(* IEC 61131-3 sources: trust-platform/crates/trust-runtime/tests/fixtures/plcopen_motion/single_axis_core/src (part 2) *)

TEST_PROGRAM plcopen_motion_single_axis_buffer_mode_support_rules_by_fb_family
VAR
    AxisHomeBuffered : AXIS_REF;
    AxisHomeUnsupported : AXIS_REF;
    AxisHaltUnsupported : AXIS_REF;
    AxisAdditiveUnsupported : AXIS_REF;
    AxisVelocityBuffered : AXIS_REF;
    AxisVelocityUnsupported : AXIS_REF;
    AxisContinuousBuffered : AXIS_REF;
    AxisContinuousUnsupported : AXIS_REF;
    SeedHomeBuffered : TRUST_MOTION_TestAxisSeed;
    SeedHomeUnsupported : TRUST_MOTION_TestAxisSeed;
    SeedHaltUnsupported : TRUST_MOTION_TestAxisSeed;
    SeedAdditiveUnsupported : TRUST_MOTION_TestAxisSeed;
    SeedVelocityBuffered : TRUST_MOTION_TestAxisSeed;
    SeedVelocityUnsupported : TRUST_MOTION_TestAxisSeed;
    SeedContinuousBuffered : TRUST_MOTION_TestAxisSeed;
    SeedContinuousUnsupported : TRUST_MOTION_TestAxisSeed;
    HomeBuffered : MC_Home;
    HomeUnsupported : MC_Home;
    HaltUnsupported : MC_Halt;
    MoveAdditiveUnsupported : MC_MoveAdditive;
    MoveVelocityBuffered : MC_MoveVelocity;
    MoveVelocityUnsupported : MC_MoveVelocity;
    MoveContinuousAbsoluteBuffered : MC_MoveContinuousAbsolute;
    MoveContinuousRelativeUnsupported : MC_MoveContinuousRelative;
END_VAR

AxisHomeBuffered.AxisId := UDINT#139;
AxisHomeBuffered.InternalIndex := UINT#18;
SeedHomeBuffered(Axis := AxisHomeBuffered, ResetDefaults := TRUE, ApplyState := TRUE, State := MC_AXIS_STATUS#mcStandstill);
HomeBuffered(Axis := AxisHomeBuffered, Execute := TRUE, Position := REAL#5.0, BufferMode := MC_BUFFER_MODE#mcBuffered);
ASSERT_TRUE(HomeBuffered.Busy);
ASSERT_TRUE(HomeBuffered.Active);
ASSERT_FALSE(HomeBuffered.Error);

AxisHomeUnsupported.AxisId := UDINT#140;
AxisHomeUnsupported.InternalIndex := UINT#19;
SeedHomeUnsupported(Axis := AxisHomeUnsupported, ResetDefaults := TRUE, ApplyState := TRUE, State := MC_AXIS_STATUS#mcStandstill);
HomeUnsupported(Axis := AxisHomeUnsupported, Execute := TRUE, Position := REAL#5.0, BufferMode := MC_BUFFER_MODE#mcBlendingLow);
ASSERT_TRUE(HomeUnsupported.Error);
ASSERT_TRUE(HomeUnsupported.ErrorID = WORD#16#0500);

AxisHaltUnsupported.AxisId := UDINT#141;
AxisHaltUnsupported.InternalIndex := UINT#20;
SeedHaltUnsupported(Axis := AxisHaltUnsupported, ResetDefaults := TRUE, ApplyState := TRUE, State := MC_AXIS_STATUS#mcContinuousMotion);
HaltUnsupported(Axis := AxisHaltUnsupported, Execute := TRUE, Deceleration := REAL#2.0, Jerk := REAL#1.0, BufferMode := MC_BUFFER_MODE#mcBlendingLow);
ASSERT_TRUE(HaltUnsupported.Error);
ASSERT_TRUE(HaltUnsupported.ErrorID = WORD#16#0500);

AxisAdditiveUnsupported.AxisId := UDINT#142;
AxisAdditiveUnsupported.InternalIndex := UINT#21;
SeedAdditiveUnsupported(
    Axis := AxisAdditiveUnsupported,
    ResetDefaults := TRUE,
    ApplyState := TRUE,
    State := MC_AXIS_STATUS#mcStandstill,
    ApplyActuals := TRUE,
    ActualPosition := REAL#10.0,
    SetPosition := REAL#10.0,
    CommandedPosition := REAL#10.0,
    ActualVelocity := REAL#0.0,
    SetVelocity := REAL#0.0,
    CommandedVelocity := REAL#0.0,
    ActualTorque := REAL#0.0
);
MoveAdditiveUnsupported(Axis := AxisAdditiveUnsupported, Execute := TRUE, ContinuousUpdate := FALSE, Distance := REAL#5.0, Velocity := REAL#4.0, Acceleration := REAL#2.0, Deceleration := REAL#2.0, Jerk := REAL#1.0, BufferMode := MC_BUFFER_MODE#mcBlendingLow);
ASSERT_TRUE(MoveAdditiveUnsupported.Error);
ASSERT_TRUE(MoveAdditiveUnsupported.ErrorID = WORD#16#0500);

AxisVelocityBuffered.AxisId := UDINT#143;
AxisVelocityBuffered.InternalIndex := UINT#22;
SeedVelocityBuffered(Axis := AxisVelocityBuffered, ResetDefaults := TRUE, ApplyState := TRUE, State := MC_AXIS_STATUS#mcStandstill);
MoveVelocityBuffered(Axis := AxisVelocityBuffered, Execute := TRUE, ContinuousUpdate := FALSE, Velocity := REAL#4.0, Acceleration := REAL#2.0, Deceleration := REAL#2.0, Jerk := REAL#1.0, Direction := MC_DIRECTION#mcCurrentDirection, BufferMode := MC_BUFFER_MODE#mcBuffered);
ASSERT_TRUE(MoveVelocityBuffered.Busy);
ASSERT_TRUE(MoveVelocityBuffered.Active);
ASSERT_TRUE(MoveVelocityBuffered.InVelocity);
ASSERT_FALSE(MoveVelocityBuffered.Error);

AxisVelocityUnsupported.AxisId := UDINT#144;
AxisVelocityUnsupported.InternalIndex := UINT#23;
SeedVelocityUnsupported(Axis := AxisVelocityUnsupported, ResetDefaults := TRUE, ApplyState := TRUE, State := MC_AXIS_STATUS#mcStandstill);
MoveVelocityUnsupported(Axis := AxisVelocityUnsupported, Execute := TRUE, ContinuousUpdate := FALSE, Velocity := REAL#4.0, Acceleration := REAL#2.0, Deceleration := REAL#2.0, Jerk := REAL#1.0, Direction := MC_DIRECTION#mcCurrentDirection, BufferMode := MC_BUFFER_MODE#mcBlendingLow);
ASSERT_TRUE(MoveVelocityUnsupported.Error);
ASSERT_TRUE(MoveVelocityUnsupported.ErrorID = WORD#16#0500);

AxisContinuousBuffered.AxisId := UDINT#145;
AxisContinuousBuffered.InternalIndex := UINT#24;
SeedContinuousBuffered(Axis := AxisContinuousBuffered, ResetDefaults := TRUE, ApplyState := TRUE, State := MC_AXIS_STATUS#mcStandstill);
MoveContinuousAbsoluteBuffered(Axis := AxisContinuousBuffered, Execute := TRUE, ContinuousUpdate := FALSE, Position := REAL#30.0, EndVelocity := REAL#3.0, Velocity := REAL#8.0, Acceleration := REAL#4.0, Deceleration := REAL#4.0, Jerk := REAL#1.0, Direction := MC_DIRECTION#mcCurrentDirection, BufferMode := MC_BUFFER_MODE#mcBuffered);
ASSERT_TRUE(MoveContinuousAbsoluteBuffered.Busy);
ASSERT_TRUE(MoveContinuousAbsoluteBuffered.Active);
ASSERT_TRUE(MoveContinuousAbsoluteBuffered.InEndVelocity);
ASSERT_FALSE(MoveContinuousAbsoluteBuffered.Error);

AxisContinuousUnsupported.AxisId := UDINT#146;
AxisContinuousUnsupported.InternalIndex := UINT#25;
SeedContinuousUnsupported(Axis := AxisContinuousUnsupported, ResetDefaults := TRUE, ApplyState := TRUE, State := MC_AXIS_STATUS#mcStandstill);
MoveContinuousRelativeUnsupported(Axis := AxisContinuousUnsupported, Execute := TRUE, ContinuousUpdate := FALSE, Distance := REAL#5.0, EndVelocity := REAL#3.0, Velocity := REAL#8.0, Acceleration := REAL#4.0, Deceleration := REAL#4.0, Jerk := REAL#1.0, BufferMode := MC_BUFFER_MODE#mcBlendingLow);
ASSERT_TRUE(MoveContinuousRelativeUnsupported.Error);
ASSERT_TRUE(MoveContinuousRelativeUnsupported.ErrorID = WORD#16#0500);
END_TEST_PROGRAM

TEST_PROGRAM plcopen_motion_single_axis_home_halt_stop_and_continuous_end_velocity_behaviors
VAR
    AxisHome : AXIS_REF;
    AxisHalt : AXIS_REF;
    AxisStop : AXIS_REF;
    AxisContinuous : AXIS_REF;
    SeedHome : TRUST_MOTION_TestAxisSeed;
    SeedHalt : TRUST_MOTION_TestAxisSeed;
    SeedStop : TRUST_MOTION_TestAxisSeed;
    SeedContinuous : TRUST_MOTION_TestAxisSeed;
    Home : MC_Home;
    Halt : MC_Halt;
    Stop : MC_Stop;
    MoveContinuousAbsolute : MC_MoveContinuousAbsolute;
    ReadStatusHome : MC_ReadStatus;
    ReadStatusHalt : MC_ReadStatus;
    ReadStatusStop : MC_ReadStatus;
    ReadStatusContinuous : MC_ReadStatus;
    ReadAxisInfo : MC_ReadAxisInfo;
    ReadActualVelocity : MC_ReadActualVelocity;
END_VAR

AxisHome.AxisId := UDINT#121;
AxisHome.InternalIndex := UINT#25;
SeedHome(Axis := AxisHome, ResetDefaults := TRUE, ApplyState := TRUE, State := MC_AXIS_STATUS#mcStandstill, ApplyPowerStage := TRUE, PowerStage := TRUE);
Home(Axis := AxisHome, Execute := TRUE, Position := REAL#12.0, BufferMode := MC_BUFFER_MODE#mcAborting);
ASSERT_TRUE(Home.Busy);
ASSERT_TRUE(Home.Active);
ReadStatusHome(Axis := AxisHome, Enable := TRUE);
ASSERT_TRUE(ReadStatusHome.Homing);
Home(Axis := AxisHome, Execute := FALSE, Position := REAL#12.0, BufferMode := MC_BUFFER_MODE#mcAborting);
ASSERT_TRUE(Home.Done);
ReadStatusHome(Axis := AxisHome, Enable := TRUE);
ASSERT_TRUE(ReadStatusHome.Standstill);
ReadAxisInfo(Axis := AxisHome, Enable := TRUE);
ASSERT_TRUE(ReadAxisInfo.IsHomed);

AxisHalt.AxisId := UDINT#122;
AxisHalt.InternalIndex := UINT#26;
SeedHalt(Axis := AxisHalt, ResetDefaults := TRUE, ApplyState := TRUE, State := MC_AXIS_STATUS#mcContinuousMotion, ApplyPowerStage := TRUE, PowerStage := TRUE);
Halt(Axis := AxisHalt, Execute := TRUE, Deceleration := REAL#2.0, Jerk := REAL#1.0, BufferMode := MC_BUFFER_MODE#mcBuffered);
ASSERT_TRUE(Halt.Busy);
ASSERT_TRUE(Halt.Active);
ReadStatusHalt(Axis := AxisHalt, Enable := TRUE);
ASSERT_TRUE(ReadStatusHalt.DiscreteMotion);
ASSERT_FALSE(ReadStatusHalt.Stopping);
Halt(Axis := AxisHalt, Execute := FALSE, Deceleration := REAL#2.0, Jerk := REAL#1.0, BufferMode := MC_BUFFER_MODE#mcBuffered);
ASSERT_TRUE(Halt.Done);
ReadStatusHalt(Axis := AxisHalt, Enable := TRUE);
ASSERT_TRUE(ReadStatusHalt.Standstill);

AxisStop.AxisId := UDINT#123;
AxisStop.InternalIndex := UINT#27;
SeedStop(Axis := AxisStop, ResetDefaults := TRUE, ApplyState := TRUE, State := MC_AXIS_STATUS#mcContinuousMotion, ApplyPowerStage := TRUE, PowerStage := TRUE);
Stop(Axis := AxisStop, Execute := TRUE, Deceleration := REAL#2.0, Jerk := REAL#1.0);
ASSERT_FALSE(Stop.Busy);
ASSERT_TRUE(Stop.Done);
ReadStatusStop(Axis := AxisStop, Enable := TRUE);
ASSERT_TRUE(ReadStatusStop.Stopping);
Stop(Axis := AxisStop, Execute := FALSE, Deceleration := REAL#2.0, Jerk := REAL#1.0);
ASSERT_TRUE(Stop.Done);
ReadStatusStop(Axis := AxisStop, Enable := TRUE);
ASSERT_TRUE(ReadStatusStop.Standstill);

AxisContinuous.AxisId := UDINT#124;
AxisContinuous.InternalIndex := UINT#28;
SeedContinuous(Axis := AxisContinuous, ResetDefaults := TRUE, ApplyState := TRUE, State := MC_AXIS_STATUS#mcStandstill);
MoveContinuousAbsolute(
    Axis := AxisContinuous,
    Execute := TRUE,
    ContinuousUpdate := FALSE,
    Position := REAL#40.0,
    EndVelocity := REAL#3.0,
    Velocity := REAL#8.0,
    Acceleration := REAL#4.0,
    Deceleration := REAL#4.0,
    Jerk := REAL#1.0,
    Direction := MC_DIRECTION#mcCurrentDirection,
    BufferMode := MC_BUFFER_MODE#mcAborting
);
ASSERT_TRUE(MoveContinuousAbsolute.Busy);
ASSERT_TRUE(MoveContinuousAbsolute.Active);
ASSERT_TRUE(MoveContinuousAbsolute.InEndVelocity);
ReadStatusContinuous(Axis := AxisContinuous, Enable := TRUE);
ASSERT_TRUE(ReadStatusContinuous.ContinuousMotion);
ReadActualVelocity(Axis := AxisContinuous, Enable := TRUE);
ASSERT_TRUE(ReadActualVelocity.Velocity = REAL#3.0);
MoveContinuousAbsolute(
    Axis := AxisContinuous,
    Execute := FALSE,
    ContinuousUpdate := FALSE,
    Position := REAL#40.0,
    EndVelocity := REAL#3.0,
    Velocity := REAL#8.0,
    Acceleration := REAL#4.0,
    Deceleration := REAL#4.0,
    Jerk := REAL#1.0,
    Direction := MC_DIRECTION#mcCurrentDirection,
    BufferMode := MC_BUFFER_MODE#mcAborting
);
ASSERT_FALSE(MoveContinuousAbsolute.InEndVelocity);
ReadStatusContinuous(Axis := AxisContinuous, Enable := TRUE);
ASSERT_TRUE(ReadStatusContinuous.Standstill);
END_TEST_PROGRAM

TEST_PROGRAM plcopen_motion_single_axis_continuous_update_changes_target_and_end_velocity
VAR
    AxisAbsolute : AXIS_REF;
    AxisRelative : AXIS_REF;
    SeedAbsolute : TRUST_MOTION_TestAxisSeed;
    SeedRelative : TRUST_MOTION_TestAxisSeed;
    MoveContinuousAbsolute : MC_MoveContinuousAbsolute;
    MoveContinuousRelative : MC_MoveContinuousRelative;
    ReadAbsolute : MC_ReadParameter;
    ReadRelative : MC_ReadParameter;
    ReadVelocityAbsolute : MC_ReadActualVelocity;
    ReadVelocityRelative : MC_ReadActualVelocity;
    Constants : MC_Constants;
END_VAR

Constants();
AxisAbsolute.AxisId := UDINT#147;
AxisAbsolute.InternalIndex := UINT#26;
SeedAbsolute(
    Axis := AxisAbsolute,
    ResetDefaults := TRUE,
    ApplyState := TRUE,
    State := MC_AXIS_STATUS#mcStandstill,
    ApplyActuals := TRUE,
    ActualPosition := REAL#10.0,
    SetPosition := REAL#10.0,
    CommandedPosition := REAL#10.0,
    ActualVelocity := REAL#0.0,
    SetVelocity := REAL#0.0,
    CommandedVelocity := REAL#0.0,
    ActualTorque := REAL#0.0
);
MoveContinuousAbsolute(Axis := AxisAbsolute, Execute := TRUE, ContinuousUpdate := FALSE, Position := REAL#40.0, EndVelocity := REAL#3.0, Velocity := REAL#8.0, Acceleration := REAL#4.0, Deceleration := REAL#4.0, Jerk := REAL#1.0, Direction := MC_DIRECTION#mcCurrentDirection, BufferMode := MC_BUFFER_MODE#mcAborting);
MoveContinuousAbsolute(Axis := AxisAbsolute, Execute := TRUE, ContinuousUpdate := TRUE, Position := REAL#55.0, EndVelocity := REAL#4.0, Velocity := REAL#8.0, Acceleration := REAL#4.0, Deceleration := REAL#4.0, Jerk := REAL#1.0, Direction := MC_DIRECTION#mcCurrentDirection, BufferMode := MC_BUFFER_MODE#mcAborting);
ASSERT_TRUE(MoveContinuousAbsolute.InEndVelocity);
ReadAbsolute(Axis := AxisAbsolute, Enable := TRUE, ParameterNumber := Constants.PN_CommandedPosition);
ASSERT_TRUE(ReadAbsolute.Value = REAL#55.0);
ReadVelocityAbsolute(Axis := AxisAbsolute, Enable := TRUE);
ASSERT_TRUE(ReadVelocityAbsolute.Velocity = REAL#4.0);

AxisRelative.AxisId := UDINT#148;
AxisRelative.InternalIndex := UINT#27;
SeedRelative(
    Axis := AxisRelative,
    ResetDefaults := TRUE,
    ApplyState := TRUE,
    State := MC_AXIS_STATUS#mcStandstill,
    ApplyActuals := TRUE,
    ActualPosition := REAL#10.0,
    SetPosition := REAL#10.0,
    CommandedPosition := REAL#10.0,
    ActualVelocity := REAL#0.0,
    SetVelocity := REAL#0.0,
    CommandedVelocity := REAL#0.0,
    ActualTorque := REAL#0.0
);
MoveContinuousRelative(Axis := AxisRelative, Execute := TRUE, ContinuousUpdate := FALSE, Distance := REAL#5.0, EndVelocity := REAL#2.0, Velocity := REAL#8.0, Acceleration := REAL#4.0, Deceleration := REAL#4.0, Jerk := REAL#1.0, BufferMode := MC_BUFFER_MODE#mcAborting);
MoveContinuousRelative(Axis := AxisRelative, Execute := TRUE, ContinuousUpdate := TRUE, Distance := REAL#8.0, EndVelocity := REAL#4.0, Velocity := REAL#8.0, Acceleration := REAL#4.0, Deceleration := REAL#4.0, Jerk := REAL#1.0, BufferMode := MC_BUFFER_MODE#mcAborting);
ASSERT_TRUE(MoveContinuousRelative.InEndVelocity);
ReadRelative(Axis := AxisRelative, Enable := TRUE, ParameterNumber := Constants.PN_CommandedPosition);
ASSERT_TRUE(ReadRelative.Value = REAL#18.0);
ReadVelocityRelative(Axis := AxisRelative, Enable := TRUE);
ASSERT_TRUE(ReadVelocityRelative.Velocity = REAL#4.0);
END_TEST_PROGRAM

TEST_PROGRAM plcopen_motion_single_axis_continuous_commandaborted_resets_in_end_velocity
VAR
    Axis : AXIS_REF;
    Seed : TRUST_MOTION_TestAxisSeed;
    MoveContinuous : MC_MoveContinuousAbsolute;
    MoveAbort : MC_MoveAbsolute;
    ReadStatus : MC_ReadStatus;
END_VAR

Axis.AxisId := UDINT#149;
Axis.InternalIndex := UINT#28;
Seed(Axis := Axis, ResetDefaults := TRUE, ApplyState := TRUE, State := MC_AXIS_STATUS#mcStandstill);
MoveContinuous(Axis := Axis, Execute := TRUE, ContinuousUpdate := FALSE, Position := REAL#30.0, EndVelocity := REAL#3.0, Velocity := REAL#8.0, Acceleration := REAL#4.0, Deceleration := REAL#4.0, Jerk := REAL#1.0, Direction := MC_DIRECTION#mcCurrentDirection, BufferMode := MC_BUFFER_MODE#mcAborting);
ASSERT_TRUE(MoveContinuous.InEndVelocity);
MoveAbort(Axis := Axis, Execute := TRUE, ContinuousUpdate := FALSE, Position := REAL#12.0, Velocity := REAL#5.0, Acceleration := REAL#2.0, Deceleration := REAL#2.0, Jerk := REAL#1.0, Direction := MC_DIRECTION#mcCurrentDirection, BufferMode := MC_BUFFER_MODE#mcAborting);
ASSERT_TRUE(MoveAbort.Active);
MoveContinuous(Axis := Axis, Execute := TRUE, ContinuousUpdate := FALSE, Position := REAL#30.0, EndVelocity := REAL#3.0, Velocity := REAL#8.0, Acceleration := REAL#4.0, Deceleration := REAL#4.0, Jerk := REAL#1.0, Direction := MC_DIRECTION#mcCurrentDirection, BufferMode := MC_BUFFER_MODE#mcAborting);
ASSERT_TRUE(MoveContinuous.CommandAborted);
ASSERT_FALSE(MoveContinuous.InEndVelocity);
ASSERT_FALSE(MoveContinuous.Busy);
ASSERT_FALSE(MoveContinuous.Active);
ReadStatus(Axis := Axis, Enable := TRUE);
ASSERT_TRUE(ReadStatus.DiscreteMotion);
END_TEST_PROGRAM

TEST_PROGRAM plcopen_motion_single_axis_buffered_home_halt_and_additive_take_ownership_after_active_motion
VAR
    AxisHome : AXIS_REF;
    AxisHalt : AXIS_REF;
    AxisAdditive : AXIS_REF;
    SeedHome : TRUST_MOTION_TestAxisSeed;
    SeedHalt : TRUST_MOTION_TestAxisSeed;
    SeedAdditive : TRUST_MOTION_TestAxisSeed;
    MoveActiveHome : MC_MoveAbsolute;
    MoveActiveHalt : MC_MoveAbsolute;
    MoveActiveAdditive : MC_MoveAbsolute;
    Home : MC_Home;
    Halt : MC_Halt;
    MoveAdditive : MC_MoveAdditive;
    ReadStatusHome : MC_ReadStatus;
    ReadStatusHalt : MC_ReadStatus;
    ReadAxisInfoHome : MC_ReadAxisInfo;
    ReadActualAdditive : MC_ReadActualPosition;
END_VAR

AxisHome.AxisId := UDINT#150;
AxisHome.InternalIndex := UINT#29;
SeedHome(Axis := AxisHome, ResetDefaults := TRUE, ApplyState := TRUE, State := MC_AXIS_STATUS#mcStandstill);
MoveActiveHome(Axis := AxisHome, Execute := TRUE, ContinuousUpdate := FALSE, Position := REAL#15.0, Velocity := REAL#5.0, Acceleration := REAL#2.0, Deceleration := REAL#2.0, Jerk := REAL#1.0, Direction := MC_DIRECTION#mcCurrentDirection, BufferMode := MC_BUFFER_MODE#mcAborting);
Home(Axis := AxisHome, Execute := TRUE, Position := REAL#7.0, BufferMode := MC_BUFFER_MODE#mcBuffered);
ASSERT_TRUE(Home.Busy);
ASSERT_FALSE(Home.Active);
MoveActiveHome(Axis := AxisHome, Execute := FALSE, ContinuousUpdate := FALSE, Position := REAL#15.0, Velocity := REAL#5.0, Acceleration := REAL#2.0, Deceleration := REAL#2.0, Jerk := REAL#1.0, Direction := MC_DIRECTION#mcCurrentDirection, BufferMode := MC_BUFFER_MODE#mcAborting);
Home(Axis := AxisHome, Execute := TRUE, Position := REAL#7.0, BufferMode := MC_BUFFER_MODE#mcBuffered);
ASSERT_TRUE(Home.Active);
ReadStatusHome(Axis := AxisHome, Enable := TRUE);
ASSERT_TRUE(ReadStatusHome.Homing);
Home(Axis := AxisHome, Execute := FALSE, Position := REAL#7.0, BufferMode := MC_BUFFER_MODE#mcBuffered);
ASSERT_TRUE(Home.Done);
ReadAxisInfoHome(Axis := AxisHome, Enable := TRUE);
ASSERT_TRUE(ReadAxisInfoHome.IsHomed);

AxisHalt.AxisId := UDINT#151;
AxisHalt.InternalIndex := UINT#30;
SeedHalt(Axis := AxisHalt, ResetDefaults := TRUE, ApplyState := TRUE, State := MC_AXIS_STATUS#mcStandstill);
MoveActiveHalt(Axis := AxisHalt, Execute := TRUE, ContinuousUpdate := FALSE, Position := REAL#20.0, Velocity := REAL#5.0, Acceleration := REAL#2.0, Deceleration := REAL#2.0, Jerk := REAL#1.0, Direction := MC_DIRECTION#mcCurrentDirection, BufferMode := MC_BUFFER_MODE#mcAborting);
Halt(Axis := AxisHalt, Execute := TRUE, Deceleration := REAL#2.0, Jerk := REAL#1.0, BufferMode := MC_BUFFER_MODE#mcBuffered);
ASSERT_TRUE(Halt.Busy);
ASSERT_FALSE(Halt.Active);
MoveActiveHalt(Axis := AxisHalt, Execute := FALSE, ContinuousUpdate := FALSE, Position := REAL#20.0, Velocity := REAL#5.0, Acceleration := REAL#2.0, Deceleration := REAL#2.0, Jerk := REAL#1.0, Direction := MC_DIRECTION#mcCurrentDirection, BufferMode := MC_BUFFER_MODE#mcAborting);
Halt(Axis := AxisHalt, Execute := TRUE, Deceleration := REAL#2.0, Jerk := REAL#1.0, BufferMode := MC_BUFFER_MODE#mcBuffered);
ASSERT_TRUE(Halt.Active);
ReadStatusHalt(Axis := AxisHalt, Enable := TRUE);
ASSERT_TRUE(ReadStatusHalt.DiscreteMotion);
Halt(Axis := AxisHalt, Execute := FALSE, Deceleration := REAL#2.0, Jerk := REAL#1.0, BufferMode := MC_BUFFER_MODE#mcBuffered);
ASSERT_TRUE(Halt.Done);
ReadStatusHalt(Axis := AxisHalt, Enable := TRUE);
ASSERT_TRUE(ReadStatusHalt.Standstill);

AxisAdditive.AxisId := UDINT#152;
AxisAdditive.InternalIndex := UINT#31;
SeedAdditive(
    Axis := AxisAdditive,
    ResetDefaults := TRUE,
    ApplyState := TRUE,
    State := MC_AXIS_STATUS#mcStandstill,
    ApplyActuals := TRUE,
    ActualPosition := REAL#10.0,
    SetPosition := REAL#10.0,
    CommandedPosition := REAL#10.0,
    ActualVelocity := REAL#0.0,
    SetVelocity := REAL#0.0,
    CommandedVelocity := REAL#0.0,
    ActualTorque := REAL#0.0
);
MoveActiveAdditive(Axis := AxisAdditive, Execute := TRUE, ContinuousUpdate := FALSE, Position := REAL#15.0, Velocity := REAL#5.0, Acceleration := REAL#2.0, Deceleration := REAL#2.0, Jerk := REAL#1.0, Direction := MC_DIRECTION#mcCurrentDirection, BufferMode := MC_BUFFER_MODE#mcAborting);
MoveAdditive(Axis := AxisAdditive, Execute := TRUE, ContinuousUpdate := FALSE, Distance := REAL#5.0, Velocity := REAL#4.0, Acceleration := REAL#2.0, Deceleration := REAL#2.0, Jerk := REAL#1.0, BufferMode := MC_BUFFER_MODE#mcBuffered);
ASSERT_TRUE(MoveAdditive.Busy);
ASSERT_FALSE(MoveAdditive.Active);
MoveActiveAdditive(Axis := AxisAdditive, Execute := FALSE, ContinuousUpdate := FALSE, Position := REAL#15.0, Velocity := REAL#5.0, Acceleration := REAL#2.0, Deceleration := REAL#2.0, Jerk := REAL#1.0, Direction := MC_DIRECTION#mcCurrentDirection, BufferMode := MC_BUFFER_MODE#mcAborting);
MoveAdditive(Axis := AxisAdditive, Execute := TRUE, ContinuousUpdate := FALSE, Distance := REAL#5.0, Velocity := REAL#4.0, Acceleration := REAL#2.0, Deceleration := REAL#2.0, Jerk := REAL#1.0, BufferMode := MC_BUFFER_MODE#mcBuffered);
ASSERT_TRUE(MoveAdditive.Active);
MoveAdditive(Axis := AxisAdditive, Execute := FALSE, ContinuousUpdate := FALSE, Distance := REAL#5.0, Velocity := REAL#4.0, Acceleration := REAL#2.0, Deceleration := REAL#2.0, Jerk := REAL#1.0, BufferMode := MC_BUFFER_MODE#mcBuffered);
ASSERT_TRUE(MoveAdditive.Done);
ReadActualAdditive(Axis := AxisAdditive, Enable := TRUE);
ASSERT_TRUE(ReadActualAdditive.Position = REAL#20.0);
END_TEST_PROGRAM

TEST_PROGRAM plcopen_motion_single_axis_move_velocity_participates_in_abort_and_buffer_queue
VAR
    AxisAbort : AXIS_REF;
    AxisBuffered : AXIS_REF;
    SeedAbort : TRUST_MOTION_TestAxisSeed;
    SeedBuffered : TRUST_MOTION_TestAxisSeed;
    MoveVelocityAbort : MC_MoveVelocity;
    MoveAbort : MC_MoveAbsolute;
    MoveActiveBuffered : MC_MoveAbsolute;
    MoveVelocityBuffered : MC_MoveVelocity;
    ReadStatusBuffered : MC_ReadStatus;
END_VAR

AxisAbort.AxisId := UDINT#153;
AxisAbort.InternalIndex := UINT#18;
SeedAbort(Axis := AxisAbort, ResetDefaults := TRUE, ApplyState := TRUE, State := MC_AXIS_STATUS#mcStandstill);
MoveVelocityAbort(Axis := AxisAbort, Execute := TRUE, ContinuousUpdate := FALSE, Velocity := REAL#4.0, Acceleration := REAL#2.0, Deceleration := REAL#2.0, Jerk := REAL#1.0, Direction := MC_DIRECTION#mcCurrentDirection, BufferMode := MC_BUFFER_MODE#mcAborting);
ASSERT_TRUE(MoveVelocityAbort.Active);
ASSERT_TRUE(MoveVelocityAbort.InVelocity);
MoveAbort(Axis := AxisAbort, Execute := TRUE, ContinuousUpdate := FALSE, Position := REAL#12.0, Velocity := REAL#5.0, Acceleration := REAL#2.0, Deceleration := REAL#2.0, Jerk := REAL#1.0, Direction := MC_DIRECTION#mcCurrentDirection, BufferMode := MC_BUFFER_MODE#mcAborting);
ASSERT_TRUE(MoveAbort.Active);
MoveVelocityAbort(Axis := AxisAbort, Execute := TRUE, ContinuousUpdate := FALSE, Velocity := REAL#4.0, Acceleration := REAL#2.0, Deceleration := REAL#2.0, Jerk := REAL#1.0, Direction := MC_DIRECTION#mcCurrentDirection, BufferMode := MC_BUFFER_MODE#mcAborting);
ASSERT_TRUE(MoveVelocityAbort.CommandAborted);
ASSERT_FALSE(MoveVelocityAbort.InVelocity);
ASSERT_FALSE(MoveVelocityAbort.Active);

AxisBuffered.AxisId := UDINT#154;
AxisBuffered.InternalIndex := UINT#19;
SeedBuffered(Axis := AxisBuffered, ResetDefaults := TRUE, ApplyState := TRUE, State := MC_AXIS_STATUS#mcStandstill);
MoveActiveBuffered(Axis := AxisBuffered, Execute := TRUE, ContinuousUpdate := FALSE, Position := REAL#16.0, Velocity := REAL#5.0, Acceleration := REAL#2.0, Deceleration := REAL#2.0, Jerk := REAL#1.0, Direction := MC_DIRECTION#mcCurrentDirection, BufferMode := MC_BUFFER_MODE#mcAborting);
MoveVelocityBuffered(Axis := AxisBuffered, Execute := TRUE, ContinuousUpdate := FALSE, Velocity := REAL#4.0, Acceleration := REAL#2.0, Deceleration := REAL#2.0, Jerk := REAL#1.0, Direction := MC_DIRECTION#mcCurrentDirection, BufferMode := MC_BUFFER_MODE#mcBuffered);
ASSERT_TRUE(MoveVelocityBuffered.Busy);
ASSERT_FALSE(MoveVelocityBuffered.Active);
MoveActiveBuffered(Axis := AxisBuffered, Execute := FALSE, ContinuousUpdate := FALSE, Position := REAL#16.0, Velocity := REAL#5.0, Acceleration := REAL#2.0, Deceleration := REAL#2.0, Jerk := REAL#1.0, Direction := MC_DIRECTION#mcCurrentDirection, BufferMode := MC_BUFFER_MODE#mcAborting);
MoveVelocityBuffered(Axis := AxisBuffered, Execute := TRUE, ContinuousUpdate := FALSE, Velocity := REAL#4.0, Acceleration := REAL#2.0, Deceleration := REAL#2.0, Jerk := REAL#1.0, Direction := MC_DIRECTION#mcCurrentDirection, BufferMode := MC_BUFFER_MODE#mcBuffered);
ASSERT_TRUE(MoveVelocityBuffered.Active);
ASSERT_TRUE(MoveVelocityBuffered.InVelocity);
ReadStatusBuffered(Axis := AxisBuffered, Enable := TRUE);
ASSERT_TRUE(ReadStatusBuffered.ContinuousMotion);
END_TEST_PROGRAM

TEST_PROGRAM plcopen_motion_single_axis_software_limits_clamp_position_target_commands
VAR
    AxisAbsoluteClamped : AXIS_REF;
    AxisRelativeClamped : AXIS_REF;
    AxisLimitDisabled : AXIS_REF;
    SeedAbsolute : TRUST_MOTION_TestAxisSeed;
    SeedRelative : TRUST_MOTION_TestAxisSeed;
    SeedDisabled : TRUST_MOTION_TestAxisSeed;
    Constants : MC_Constants;
    WriteParameterAbsolute : MC_WriteParameter;
    WriteBoolAbsolute : MC_WriteBoolParameter;
    MoveAbsolute : MC_MoveAbsolute;
    ReadActualAbsolute : MC_ReadActualPosition;
    WriteParameterRelative : MC_WriteParameter;
    WriteBoolRelative : MC_WriteBoolParameter;
    MoveRelative : MC_MoveRelative;
    ReadActualRelative : MC_ReadActualPosition;
    WriteParameterDisabled : MC_WriteParameter;
    MoveAbsoluteDisabled : MC_MoveAbsolute;
    ReadActualDisabled : MC_ReadActualPosition;
END_VAR

Constants();
AxisAbsoluteClamped.AxisId := UDINT#156;
AxisAbsoluteClamped.InternalIndex := UINT#14;
SeedAbsolute(
    Axis := AxisAbsoluteClamped,
    ResetDefaults := TRUE,
    ApplyState := TRUE,
    State := MC_AXIS_STATUS#mcStandstill,
    ApplyActuals := TRUE,
    ActualPosition := REAL#10.0,
    SetPosition := REAL#10.0,
    CommandedPosition := REAL#10.0,
    ActualVelocity := REAL#0.0,
    SetVelocity := REAL#0.0,
    CommandedVelocity := REAL#0.0,
    ActualTorque := REAL#0.0
);
WriteParameterAbsolute(Axis := AxisAbsoluteClamped, Execute := TRUE, ParameterNumber := Constants.PN_SWLimitPos, Value := REAL#25.0, ExecutionMode := MC_EXECUTION_MODE#mcImmediately);
WriteParameterAbsolute(Axis := AxisAbsoluteClamped, Execute := FALSE, ParameterNumber := Constants.PN_SWLimitPos, Value := REAL#25.0, ExecutionMode := MC_EXECUTION_MODE#mcImmediately);
WriteBoolAbsolute(Axis := AxisAbsoluteClamped, Execute := TRUE, ParameterNumber := Constants.PN_EnableLimitPos, Value := TRUE, ExecutionMode := MC_EXECUTION_MODE#mcImmediately);
WriteBoolAbsolute(Axis := AxisAbsoluteClamped, Execute := FALSE, ParameterNumber := Constants.PN_EnableLimitPos, Value := TRUE, ExecutionMode := MC_EXECUTION_MODE#mcImmediately);
MoveAbsolute(Axis := AxisAbsoluteClamped, Execute := TRUE, ContinuousUpdate := FALSE, Position := REAL#40.0, Velocity := REAL#6.0, Acceleration := REAL#2.0, Deceleration := REAL#2.0, Jerk := REAL#1.0, Direction := MC_DIRECTION#mcCurrentDirection, BufferMode := MC_BUFFER_MODE#mcAborting);
ASSERT_TRUE(MoveAbsolute.Active);
ASSERT_FALSE(MoveAbsolute.Error);
MoveAbsolute(Axis := AxisAbsoluteClamped, Execute := FALSE, ContinuousUpdate := FALSE, Position := REAL#40.0, Velocity := REAL#6.0, Acceleration := REAL#2.0, Deceleration := REAL#2.0, Jerk := REAL#1.0, Direction := MC_DIRECTION#mcCurrentDirection, BufferMode := MC_BUFFER_MODE#mcAborting);
ASSERT_TRUE(MoveAbsolute.Done);
ReadActualAbsolute(Axis := AxisAbsoluteClamped, Enable := TRUE);
ASSERT_TRUE(ReadActualAbsolute.Position = REAL#25.0);

AxisRelativeClamped.AxisId := UDINT#157;
AxisRelativeClamped.InternalIndex := UINT#15;
SeedRelative(
    Axis := AxisRelativeClamped,
    ResetDefaults := TRUE,
    ApplyState := TRUE,
    State := MC_AXIS_STATUS#mcStandstill,
    ApplyActuals := TRUE,
    ActualPosition := REAL#10.0,
    SetPosition := REAL#10.0,
    CommandedPosition := REAL#10.0,
    ActualVelocity := REAL#0.0,
    SetVelocity := REAL#0.0,
    CommandedVelocity := REAL#0.0,
    ActualTorque := REAL#0.0
);
WriteParameterRelative(Axis := AxisRelativeClamped, Execute := TRUE, ParameterNumber := Constants.PN_SWLimitNeg, Value := REAL#0.0 - REAL#5.0, ExecutionMode := MC_EXECUTION_MODE#mcImmediately);
WriteParameterRelative(Axis := AxisRelativeClamped, Execute := FALSE, ParameterNumber := Constants.PN_SWLimitNeg, Value := REAL#0.0 - REAL#5.0, ExecutionMode := MC_EXECUTION_MODE#mcImmediately);
WriteBoolRelative(Axis := AxisRelativeClamped, Execute := TRUE, ParameterNumber := Constants.PN_EnableLimitNeg, Value := TRUE, ExecutionMode := MC_EXECUTION_MODE#mcImmediately);
WriteBoolRelative(Axis := AxisRelativeClamped, Execute := FALSE, ParameterNumber := Constants.PN_EnableLimitNeg, Value := TRUE, ExecutionMode := MC_EXECUTION_MODE#mcImmediately);
MoveRelative(Axis := AxisRelativeClamped, Execute := TRUE, ContinuousUpdate := FALSE, Distance := REAL#0.0 - REAL#30.0, Velocity := REAL#6.0, Acceleration := REAL#2.0, Deceleration := REAL#2.0, Jerk := REAL#1.0, BufferMode := MC_BUFFER_MODE#mcAborting);
ASSERT_TRUE(MoveRelative.Active);
ASSERT_FALSE(MoveRelative.Error);
MoveRelative(Axis := AxisRelativeClamped, Execute := FALSE, ContinuousUpdate := FALSE, Distance := REAL#0.0 - REAL#30.0, Velocity := REAL#6.0, Acceleration := REAL#2.0, Deceleration := REAL#2.0, Jerk := REAL#1.0, BufferMode := MC_BUFFER_MODE#mcAborting);
ASSERT_TRUE(MoveRelative.Done);
ReadActualRelative(Axis := AxisRelativeClamped, Enable := TRUE);
ASSERT_TRUE(ReadActualRelative.Position = REAL#0.0 - REAL#5.0);

AxisLimitDisabled.AxisId := UDINT#158;
AxisLimitDisabled.InternalIndex := UINT#16;
SeedDisabled(
    Axis := AxisLimitDisabled,
    ResetDefaults := TRUE,
    ApplyState := TRUE,
    State := MC_AXIS_STATUS#mcStandstill,
    ApplyActuals := TRUE,
    ActualPosition := REAL#10.0,
    SetPosition := REAL#10.0,
    CommandedPosition := REAL#10.0,
    ActualVelocity := REAL#0.0,
    SetVelocity := REAL#0.0,
    CommandedVelocity := REAL#0.0,
    ActualTorque := REAL#0.0
);
WriteParameterDisabled(Axis := AxisLimitDisabled, Execute := TRUE, ParameterNumber := Constants.PN_SWLimitPos, Value := REAL#25.0, ExecutionMode := MC_EXECUTION_MODE#mcImmediately);
WriteParameterDisabled(Axis := AxisLimitDisabled, Execute := FALSE, ParameterNumber := Constants.PN_SWLimitPos, Value := REAL#25.0, ExecutionMode := MC_EXECUTION_MODE#mcImmediately);
MoveAbsoluteDisabled(Axis := AxisLimitDisabled, Execute := TRUE, ContinuousUpdate := FALSE, Position := REAL#40.0, Velocity := REAL#6.0, Acceleration := REAL#2.0, Deceleration := REAL#2.0, Jerk := REAL#1.0, Direction := MC_DIRECTION#mcCurrentDirection, BufferMode := MC_BUFFER_MODE#mcAborting);
ASSERT_TRUE(MoveAbsoluteDisabled.Active);
ASSERT_FALSE(MoveAbsoluteDisabled.Error);
MoveAbsoluteDisabled(Axis := AxisLimitDisabled, Execute := FALSE, ContinuousUpdate := FALSE, Position := REAL#40.0, Velocity := REAL#6.0, Acceleration := REAL#2.0, Deceleration := REAL#2.0, Jerk := REAL#1.0, Direction := MC_DIRECTION#mcCurrentDirection, BufferMode := MC_BUFFER_MODE#mcAborting);
ASSERT_TRUE(MoveAbsoluteDisabled.Done);
ReadActualDisabled(Axis := AxisLimitDisabled, Enable := TRUE);
ASSERT_TRUE(ReadActualDisabled.Position = REAL#40.0);
END_TEST_PROGRAM

TEST_PROGRAM plcopen_motion_single_axis_move_absolute_final_position_semantics
VAR
    Axis : AXIS_REF;
    Seed : TRUST_MOTION_TestAxisSeed;
    MoveAbsolute : MC_MoveAbsolute;
    ReadActualPosition : MC_ReadActualPosition;
END_VAR

Axis.AxisId := UDINT#125;
Axis.InternalIndex := UINT#29;
Seed(
    Axis := Axis,
    ResetDefaults := TRUE,
    ApplyState := TRUE,
    State := MC_AXIS_STATUS#mcStandstill,
    ApplyActuals := TRUE,
    ActualPosition := REAL#10.0,
    SetPosition := REAL#10.0,
    CommandedPosition := REAL#10.0,
    ActualVelocity := REAL#0.0,
    SetVelocity := REAL#0.0,
    CommandedVelocity := REAL#0.0,
    ActualTorque := REAL#0.0
);
MoveAbsolute(
    Axis := Axis,
    Execute := TRUE,
    ContinuousUpdate := FALSE,
    Position := REAL#42.0,
    Velocity := REAL#8.0,
    Acceleration := REAL#4.0,
    Deceleration := REAL#4.0,
    Jerk := REAL#1.0,
    Direction := MC_DIRECTION#mcCurrentDirection,
    BufferMode := MC_BUFFER_MODE#mcAborting
);
ASSERT_TRUE(MoveAbsolute.Busy);
ASSERT_TRUE(MoveAbsolute.Active);
ASSERT_FALSE(MoveAbsolute.Done);
MoveAbsolute(
    Axis := Axis,
    Execute := FALSE,
    ContinuousUpdate := FALSE,
    Position := REAL#42.0,
    Velocity := REAL#8.0,
    Acceleration := REAL#4.0,
    Deceleration := REAL#4.0,
    Jerk := REAL#1.0,
    Direction := MC_DIRECTION#mcCurrentDirection,
    BufferMode := MC_BUFFER_MODE#mcAborting
);
ASSERT_TRUE(MoveAbsolute.Done);
ReadActualPosition(Axis := Axis, Enable := TRUE);
ASSERT_TRUE(ReadActualPosition.Position = REAL#42.0);
END_TEST_PROGRAM

TEST_PROGRAM plcopen_motion_single_axis_home_from_nonstandstill_entry_state
VAR
    Axis : AXIS_REF;
    Seed : TRUST_MOTION_TestAxisSeed;
    Home : MC_Home;
    ReadStatus : MC_ReadStatus;
END_VAR

Axis.AxisId := UDINT#126;
Axis.InternalIndex := UINT#30;
Seed(Axis := Axis, ResetDefaults := TRUE, ApplyState := TRUE, State := MC_AXIS_STATUS#mcDiscreteMotion, ApplyPowerStage := TRUE, PowerStage := TRUE);
Home(Axis := Axis, Execute := TRUE, Position := REAL#5.0, BufferMode := MC_BUFFER_MODE#mcAborting);
ASSERT_TRUE(Home.Busy);
ASSERT_TRUE(Home.Active);
ASSERT_FALSE(Home.Error);
ReadStatus(Axis := Axis, Enable := TRUE);
ASSERT_TRUE(ReadStatus.Homing);
Home(Axis := Axis, Execute := FALSE, Position := REAL#5.0, BufferMode := MC_BUFFER_MODE#mcAborting);
ASSERT_TRUE(Home.Done);
ReadStatus(Axis := Axis, Enable := TRUE);
ASSERT_TRUE(ReadStatus.Standstill);
END_TEST_PROGRAM

TEST_PROGRAM plcopen_motion_single_axis_end_to_end_conformance_scenario
VAR
    AxisPowerMotion : AXIS_REF;
    AxisHaltStop : AXIS_REF;
    AxisFaultReset : AXIS_REF;
    SeedPowerMotion : TRUST_MOTION_TestAxisSeed;
    SeedHaltStop : TRUST_MOTION_TestAxisSeed;
    SeedFaultReset : TRUST_MOTION_TestAxisSeed;
    Constants : MC_Constants;
    PowerPowerMotion : MC_Power;
    WriteParameterPowerMotion : MC_WriteParameter;
    WriteBoolPowerMotion : MC_WriteBoolParameter;
    MoveAbsolutePowerMotion : MC_MoveAbsolute;
    ReadStatusPowerMotion : MC_ReadStatus;
    ReadActualPositionPowerMotion : MC_ReadActualPosition;
    MoveVelocityHalt : MC_MoveVelocity;
    MoveVelocityStop : MC_MoveVelocity;
    HaltHaltStop : MC_Halt;
    StopHaltStop : MC_Stop;
    ReadStatusHaltStop : MC_ReadStatus;
    MoveAbsoluteFaultReset : MC_MoveAbsolute;
    ReadStatusFaultReset : MC_ReadStatus;
    ReadAxisErrorFaultReset : MC_ReadAxisError;
    ResetFaultReset : MC_Reset;
END_VAR

Constants();

AxisPowerMotion.AxisId := UDINT#159;
AxisPowerMotion.InternalIndex := UINT#17;
SeedPowerMotion(
    Axis := AxisPowerMotion,
    ResetDefaults := TRUE,
    ApplyState := TRUE,
    State := MC_AXIS_STATUS#mcDisabled,
    ApplyPowerStage := TRUE,
    PowerStage := FALSE,
    ApplyActuals := TRUE,
    ActualPosition := REAL#10.0,
    SetPosition := REAL#10.0,
    CommandedPosition := REAL#10.0,
    ActualVelocity := REAL#0.0,
    SetVelocity := REAL#0.0,
    CommandedVelocity := REAL#0.0,
    ActualTorque := REAL#0.0
);
PowerPowerMotion(Axis := AxisPowerMotion, Enable := TRUE);
ASSERT_TRUE(PowerPowerMotion.Status);
ReadStatusPowerMotion(Axis := AxisPowerMotion, Enable := TRUE);
ASSERT_TRUE(ReadStatusPowerMotion.Standstill);
WriteParameterPowerMotion(Axis := AxisPowerMotion, Execute := TRUE, ParameterNumber := Constants.PN_MaxVelocityAppl, Value := REAL#8.0, ExecutionMode := MC_EXECUTION_MODE#mcImmediately);
ASSERT_TRUE(WriteParameterPowerMotion.Done);
WriteParameterPowerMotion(Axis := AxisPowerMotion, Execute := FALSE, ParameterNumber := Constants.PN_MaxVelocityAppl, Value := REAL#8.0, ExecutionMode := MC_EXECUTION_MODE#mcImmediately);
WriteParameterPowerMotion(Axis := AxisPowerMotion, Execute := TRUE, ParameterNumber := Constants.PN_SWLimitPos, Value := REAL#30.0, ExecutionMode := MC_EXECUTION_MODE#mcImmediately);
ASSERT_TRUE(WriteParameterPowerMotion.Done);
WriteParameterPowerMotion(Axis := AxisPowerMotion, Execute := FALSE, ParameterNumber := Constants.PN_SWLimitPos, Value := REAL#30.0, ExecutionMode := MC_EXECUTION_MODE#mcImmediately);
WriteBoolPowerMotion(Axis := AxisPowerMotion, Execute := TRUE, ParameterNumber := Constants.PN_EnableLimitPos, Value := TRUE, ExecutionMode := MC_EXECUTION_MODE#mcImmediately);
ASSERT_TRUE(WriteBoolPowerMotion.Done);
WriteBoolPowerMotion(Axis := AxisPowerMotion, Execute := FALSE, ParameterNumber := Constants.PN_EnableLimitPos, Value := TRUE, ExecutionMode := MC_EXECUTION_MODE#mcImmediately);
MoveAbsolutePowerMotion(Axis := AxisPowerMotion, Execute := TRUE, ContinuousUpdate := FALSE, Position := REAL#40.0, Velocity := REAL#8.0, Acceleration := REAL#2.0, Deceleration := REAL#2.0, Jerk := REAL#1.0, Direction := MC_DIRECTION#mcCurrentDirection, BufferMode := MC_BUFFER_MODE#mcAborting);
ASSERT_TRUE(MoveAbsolutePowerMotion.Active);
MoveAbsolutePowerMotion(Axis := AxisPowerMotion, Execute := FALSE, ContinuousUpdate := FALSE, Position := REAL#40.0, Velocity := REAL#8.0, Acceleration := REAL#2.0, Deceleration := REAL#2.0, Jerk := REAL#1.0, Direction := MC_DIRECTION#mcCurrentDirection, BufferMode := MC_BUFFER_MODE#mcAborting);
ASSERT_TRUE(MoveAbsolutePowerMotion.Done);
ReadActualPositionPowerMotion(Axis := AxisPowerMotion, Enable := TRUE);
ASSERT_TRUE(ReadActualPositionPowerMotion.Position = REAL#30.0);

AxisHaltStop.AxisId := UDINT#160;
AxisHaltStop.InternalIndex := UINT#18;
SeedHaltStop(Axis := AxisHaltStop, ResetDefaults := TRUE, ApplyState := TRUE, State := MC_AXIS_STATUS#mcStandstill, ApplyPowerStage := TRUE, PowerStage := TRUE);
MoveVelocityHalt(Axis := AxisHaltStop, Execute := TRUE, ContinuousUpdate := FALSE, Velocity := REAL#4.0, Acceleration := REAL#2.0, Deceleration := REAL#2.0, Jerk := REAL#1.0, Direction := MC_DIRECTION#mcCurrentDirection, BufferMode := MC_BUFFER_MODE#mcAborting);
ASSERT_TRUE(MoveVelocityHalt.InVelocity);
HaltHaltStop(Axis := AxisHaltStop, Execute := TRUE, Deceleration := REAL#2.0, Jerk := REAL#1.0, BufferMode := MC_BUFFER_MODE#mcAborting);
ASSERT_TRUE(HaltHaltStop.Active);
HaltHaltStop(Axis := AxisHaltStop, Execute := FALSE, Deceleration := REAL#2.0, Jerk := REAL#1.0, BufferMode := MC_BUFFER_MODE#mcAborting);
ASSERT_TRUE(HaltHaltStop.Done);
ReadStatusHaltStop(Axis := AxisHaltStop, Enable := TRUE);
ASSERT_TRUE(ReadStatusHaltStop.Standstill);
MoveVelocityStop(Axis := AxisHaltStop, Execute := TRUE, ContinuousUpdate := FALSE, Velocity := REAL#3.0, Acceleration := REAL#2.0, Deceleration := REAL#2.0, Jerk := REAL#1.0, Direction := MC_DIRECTION#mcCurrentDirection, BufferMode := MC_BUFFER_MODE#mcAborting);
ASSERT_TRUE(MoveVelocityStop.InVelocity);
StopHaltStop(Axis := AxisHaltStop, Execute := TRUE, Deceleration := REAL#2.0, Jerk := REAL#1.0);
ASSERT_FALSE(StopHaltStop.Busy);
ASSERT_TRUE(StopHaltStop.Done);
ReadStatusHaltStop(Axis := AxisHaltStop, Enable := TRUE);
ASSERT_TRUE(ReadStatusHaltStop.Stopping);
StopHaltStop(Axis := AxisHaltStop, Execute := FALSE, Deceleration := REAL#2.0, Jerk := REAL#1.0);
ReadStatusHaltStop(Axis := AxisHaltStop, Enable := TRUE);
ASSERT_TRUE(ReadStatusHaltStop.Standstill);

AxisFaultReset.AxisId := UDINT#161;
AxisFaultReset.InternalIndex := UINT#19;
SeedFaultReset(Axis := AxisFaultReset, ResetDefaults := TRUE, ApplyState := TRUE, State := MC_AXIS_STATUS#mcStandstill, ApplyPowerStage := TRUE, PowerStage := TRUE);
MoveAbsoluteFaultReset(Axis := AxisFaultReset, Execute := TRUE, ContinuousUpdate := FALSE, Position := REAL#22.0, Velocity := REAL#6.0, Acceleration := REAL#2.0, Deceleration := REAL#2.0, Jerk := REAL#1.0, Direction := MC_DIRECTION#mcCurrentDirection, BufferMode := MC_BUFFER_MODE#mcAborting);
ASSERT_TRUE(MoveAbsoluteFaultReset.Active);
SeedFaultReset(Axis := AxisFaultReset, ResetDefaults := FALSE, ApplyState := FALSE, ApplyPowerStage := FALSE, ApplyAxisError := TRUE, AxisErrorID := WORD#16#0200);
MoveAbsoluteFaultReset(Axis := AxisFaultReset, Execute := TRUE, ContinuousUpdate := FALSE, Position := REAL#22.0, Velocity := REAL#6.0, Acceleration := REAL#2.0, Deceleration := REAL#2.0, Jerk := REAL#1.0, Direction := MC_DIRECTION#mcCurrentDirection, BufferMode := MC_BUFFER_MODE#mcAborting);
ASSERT_TRUE(MoveAbsoluteFaultReset.Error);
ASSERT_TRUE(MoveAbsoluteFaultReset.ErrorID = WORD#16#0200);
ReadStatusFaultReset(Axis := AxisFaultReset, Enable := TRUE);
ASSERT_TRUE(ReadStatusFaultReset.ErrorStop);
ReadAxisErrorFaultReset(Axis := AxisFaultReset, Enable := TRUE);
ASSERT_TRUE(ReadAxisErrorFaultReset.Valid);
ASSERT_TRUE(ReadAxisErrorFaultReset.AxisErrorID = WORD#16#0200);
ResetFaultReset(Axis := AxisFaultReset, Execute := TRUE);
ASSERT_TRUE(ResetFaultReset.Done);
ResetFaultReset(Axis := AxisFaultReset, Execute := FALSE);
ReadStatusFaultReset(Axis := AxisFaultReset, Enable := TRUE);
ASSERT_TRUE(ReadStatusFaultReset.Standstill);
END_TEST_PROGRAM

TEST_PROGRAM plcopen_motion_single_axis_dynamic_max_parameter_rejections
VAR
    Axis : AXIS_REF;
    Constants : MC_Constants;
    WriteParameter : MC_WriteParameter;
END_VAR

Axis.AxisId := UDINT#127;
Axis.InternalIndex := UINT#31;
Constants();
WriteParameter(Axis := Axis, Execute := TRUE, ParameterNumber := Constants.PN_MaxVelocityAppl, Value := REAL#0.0, ExecutionMode := MC_EXECUTION_MODE#mcImmediately);
ASSERT_TRUE(WriteParameter.Error);
ASSERT_TRUE(WriteParameter.ErrorID = WORD#16#0001);
WriteParameter(Axis := Axis, Execute := FALSE, ParameterNumber := Constants.PN_MaxVelocityAppl, Value := REAL#0.0, ExecutionMode := MC_EXECUTION_MODE#mcImmediately);
WriteParameter(Axis := Axis, Execute := TRUE, ParameterNumber := Constants.PN_MaxAccelerationAppl, Value := REAL#0.0 - REAL#1.0, ExecutionMode := MC_EXECUTION_MODE#mcImmediately);
ASSERT_TRUE(WriteParameter.Error);
ASSERT_TRUE(WriteParameter.ErrorID = WORD#16#0001);
WriteParameter(Axis := Axis, Execute := FALSE, ParameterNumber := Constants.PN_MaxAccelerationAppl, Value := REAL#0.0 - REAL#1.0, ExecutionMode := MC_EXECUTION_MODE#mcImmediately);
WriteParameter(Axis := Axis, Execute := TRUE, ParameterNumber := Constants.PN_MaxDecelerationAppl, Value := REAL#0.0, ExecutionMode := MC_EXECUTION_MODE#mcImmediately);
ASSERT_TRUE(WriteParameter.Error);
ASSERT_TRUE(WriteParameter.ErrorID = WORD#16#0001);
WriteParameter(Axis := Axis, Execute := FALSE, ParameterNumber := Constants.PN_MaxDecelerationAppl, Value := REAL#0.0, ExecutionMode := MC_EXECUTION_MODE#mcImmediately);
WriteParameter(Axis := Axis, Execute := TRUE, ParameterNumber := Constants.PN_MaxJerkAppl, Value := REAL#0.0 - REAL#1.0, ExecutionMode := MC_EXECUTION_MODE#mcImmediately);
ASSERT_TRUE(WriteParameter.Error);
ASSERT_TRUE(WriteParameter.ErrorID = WORD#16#0001);
WriteParameter(Axis := Axis, Execute := FALSE, ParameterNumber := Constants.PN_MaxJerkAppl, Value := REAL#0.0 - REAL#1.0, ExecutionMode := MC_EXECUTION_MODE#mcImmediately);
END_TEST_PROGRAM
